// ---- POUs/err.TcPOU
FUNCTION_BLOCK err
VAR_INPUT
	enter : BOOL;
END_VAR
VAR_OUTPUT
END_VAR
VAR
	i:INT;
	step:INT:=0;
	pulse_timer:TON;
	retry_timer:TON;
	has_err:BOOL;
	has_power_not_ready:BOOL;
	has_other_error:BOOL;
	all_powered:BOOL;
	backoff_move : ARRAY[1..7] OF MC_MoveRelative;
	backoff_exec : ARRAY[1..7] OF BOOL;
	backoff_distance : ARRAY[1..7] OF LREAL;
	backoff_attempts : ARRAY[1..7] OF UINT;
	backoff_blocked : BOOL;
	backoff_needed : BOOL;
	backoff_finished : BOOL;
	backoff_error : BOOL;
	backoff_disabled : BOOL;
	power_not_ready_errid : UDINT := 16#00004650;
END_VAR

(* 
Error recovery state:
  - disable external setpoint generation and keep estop hold active
  - if the only active power error is 16#00004650, recover by cycling MC_Power.Enable
  - other errors still use MC_Reset
  - leave _err only after errors are gone and all axes are powered again
*)

has_err := FALSE;
has_power_not_ready := FALSE;
has_other_error := FALSE;
all_powered := TRUE;

FOR i:=1 TO 7 DO
	IF NOT G.power_output[i].Done THEN
		all_powered := FALSE;
	END_IF

	IF G.axis[i].Status.Error OR G.axis[i].Status.DriveDeviceError OR G.power_output[i].Error OR G.reset_output[i].Error THEN
		has_err := TRUE;

		IF (G.power_output[i].Error AND (G.power_output[i].ErrorID = power_not_ready_errid))
		   OR (G.axis[i].Status.Error AND (G.axis[i].Status.ErrorID = power_not_ready_errid)) THEN
			has_power_not_ready := TRUE;
		END_IF

		IF (G.axis[i].Status.Error AND (G.axis[i].Status.ErrorID <> power_not_ready_errid))
		   OR G.axis[i].Status.DriveDeviceError
		   OR G.reset_output[i].Error
		   OR (G.power_output[i].Error AND (G.power_output[i].ErrorID <> power_not_ready_errid)) THEN
			has_other_error := TRUE;
		END_IF
	END_IF
END_FOR

G.estop_hold_req := TRUE;
IF enter THEN
	FOR i:=1 TO 7 DO
		backoff_attempts[i] := 0;
		backoff_exec[i] := FALSE;
		G.err_backoff_failed[i] := FALSE;
		G.err_backoff_active[i] := FALSE;
	END_FOR
END_IF
FOR i:=1 TO 7 DO
	backoff_move[i](Axis:=G.axis[i], Execute:=backoff_exec[i],
		Distance:=backoff_distance[i], Velocity:=G.err_backoff_velocity,
		Acceleration:=G.err_backoff_acc, Deceleration:=G.err_backoff_acc);
END_FOR
backoff_blocked := FALSE;
backoff_needed := FALSE;
IF G.self_check_done AND ((step = 1) OR (step = 3) OR (step = 11)) AND NOT has_err AND all_powered THEN
	backoff_disabled := TRUE;
	FOR i:=1 TO 7 DO
		IF ((i = 1) OR (i = 3) OR (i = 5) OR (i = 6)) AND G.axis[i].Status.DriveLimitActive
			AND G.SetPointGenDisable[i].Enabled THEN backoff_disabled := FALSE; END_IF
	END_FOR
	IF NOT backoff_disabled THEN
		FOR i:=1 TO 7 DO
			G.SetPointGenEnable[i].Execute := FALSE;
			G.SetPointGenDisable[i].Execute := TRUE;
		END_FOR
		RETURN;
	END_IF
	FOR i:=1 TO 7 DO
		IF ((i = 1) OR (i = 3) OR (i = 5) OR (i = 6)) AND G.axis[i].Status.DriveLimitActive THEN
			backoff_blocked := TRUE;
			IF backoff_attempts[i] < G.recovery_max_retries THEN
				IF G.axis[i].NcToPlc.ActPos - G.leftlimit[i] <=
					G.leftlimit[i] + G.rslimit_distance[i] - G.axis[i].NcToPlc.ActPos THEN
					backoff_distance[i] := G.err_backoff_distance;
				ELSE
					backoff_distance[i] := -G.err_backoff_distance;
				END_IF
				backoff_attempts[i] := backoff_attempts[i] + 1;
				backoff_exec[i] := TRUE;
				G.err_backoff_active[i] := TRUE;
				backoff_needed := TRUE;
			ELSE
				G.err_backoff_failed[i] := TRUE;
			END_IF
		END_IF
	END_FOR
	IF backoff_needed THEN step := 20; END_IF
END_IF
IF step = 20 THEN
	backoff_finished := TRUE;
	backoff_error := has_err;
	FOR i:=1 TO 7 DO
		G.SetPointGenEnable[i].Execute := FALSE;
		G.SetPointGenDisable[i].Execute := TRUE;
		IF G.err_backoff_active[i] THEN
			IF backoff_move[i].Error OR backoff_move[i].CommandAborted THEN
				backoff_error := TRUE;
			ELSIF NOT backoff_move[i].Done THEN
				backoff_finished := FALSE;
			END_IF
		END_IF
	END_FOR
	IF backoff_error OR backoff_finished THEN
		FOR i:=1 TO 7 DO
			backoff_exec[i] := FALSE;
			G.err_backoff_active[i] := FALSE;
		END_FOR
		// 重置流程提供下降沿；仍压限位时按本次进入err的剩余次数再退离。
		step := 0;
	END_IF
	RETURN;
END_IF

CASE step OF
0:
	FOR i:=1 TO 7 DO
		G.SetPointGenEnable[i].Execute := FALSE;
		G.SetPointGenDisable[i].Execute := TRUE;
		G.axis_Reset[i].Execute := FALSE;
	END_FOR
	pulse_timer(IN:=FALSE);
	retry_timer(IN:=FALSE);
	step := 1;

1:
	FOR i:=1 TO 7 DO
		G.SetPointGenDisable[i].Execute := FALSE;
	END_FOR

	IF (NOT has_err) AND all_powered AND NOT backoff_blocked THEN
		step := 0;
		G.gen_state := _clear_err;
		RETURN;
	END_IF

	IF NOT has_err THEN
		FOR i:=1 TO 7 DO
			G.axis_Reset[i].Execute := FALSE;
			G.power_[i].Enable := FALSE;
		END_FOR
		pulse_timer(IN:=TRUE, PT:=T#200MS);
		step := 10;
		RETURN;
	END_IF

	IF has_power_not_ready AND NOT has_other_error THEN
		pulse_timer(IN:=TRUE, PT:=T#200MS);
		retry_timer(IN:=FALSE);
		step := 10;
		RETURN;
	END_IF

	FOR i:=1 TO 7 DO
		IF G.axis[i].Status.Error OR G.axis[i].Status.DriveDeviceError OR G.power_output[i].Error OR G.reset_output[i].Error THEN
			G.axis_Reset[i].Execute := TRUE;
		END_IF
	END_FOR
	pulse_timer(IN:=TRUE, PT:=T#200MS);
	step := 2;

2:
	pulse_timer(IN:=TRUE);
	IF pulse_timer.Q THEN
		FOR i:=1 TO 7 DO
			G.axis_Reset[i].Execute := FALSE;
		END_FOR
		pulse_timer(IN:=FALSE);
		retry_timer(IN:=TRUE, PT:=T#2S);
		step := 3;
	END_IF

3:
	retry_timer(IN:=TRUE);

	IF (NOT has_err) AND all_powered AND NOT backoff_blocked THEN
		retry_timer(IN:=FALSE);
		step := 0;
		G.gen_state := _clear_err;
		RETURN;
	END_IF

	IF retry_timer.Q THEN
		retry_timer(IN:=FALSE);
		step := 1;
	END_IF

10:
	FOR i:=1 TO 7 DO
		IF (G.power_output[i].Error AND (G.power_output[i].ErrorID = power_not_ready_errid))
		   OR (G.axis[i].Status.Error AND (G.axis[i].Status.ErrorID = power_not_ready_errid))
		   OR G.axis[i].Status.DriveDeviceError THEN
			G.power_[i].Enable := FALSE;
			G.axis_Reset[i].Execute := TRUE;
		ELSE
			G.power_[i].Enable := TRUE;
			G.axis_Reset[i].Execute := FALSE;
		END_IF
	END_FOR

	pulse_timer(IN:=TRUE, PT:=T#200MS);
	IF pulse_timer.Q THEN
		pulse_timer(IN:=FALSE);
		FOR i:=1 TO 7 DO
			G.axis_Reset[i].Execute := FALSE;
			G.power_[i].Enable := TRUE;
		END_FOR
		retry_timer(IN:=TRUE, PT:=T#3S);
		step := 11;
	END_IF

11:
	FOR i:=1 TO 7 DO
		G.power_[i].Enable := TRUE;
	END_FOR

	retry_timer(IN:=TRUE);

	IF (NOT has_err) AND all_powered AND NOT backoff_blocked THEN
		retry_timer(IN:=FALSE);
		step := 0;
		G.gen_state := _clear_err;
		RETURN;
	END_IF

	IF has_err THEN
		retry_timer(IN:=FALSE);
		step := 1;
		RETURN;
	END_IF

	IF retry_timer.Q THEN
		retry_timer(IN:=FALSE);
		step := 1;
	END_IF
END_CASE

END_FUNCTION_BLOCK

// ---- POUs/reset.TcPOU
FUNCTION_BLOCK reset
VAR_INPUT
END_VAR
VAR_OUTPUT
END_VAR
VAR
	i:INT;
	step:INT:=0;
	reset_timer:TON;
	all_done:BOOL;
END_VAR

(*
FUNCTION_BLOCK: reset
功能说明:
  故障复位流程：对错误轴发出 MC_Reset 清错请求，清错后回到 _init；若错误仍在则转入 _err。

状态机(step):
  0) 预处理：拉低 Execute 形成上升沿；同时请求禁用外部给定模式(避免复位期间被 refer 干预)
  1) 触发复位：对 7 轴发出 MC_Reset.Execute=TRUE，并启动超时计时器
  2) 等待：Done/Error/错误已清除 或超时则收尾并决定跳转(_init/_err)
*)

CASE step OF
0:
	// 预处理：确保后续有上升沿，同时在复位阶段禁用外部给定
	FOR i:=1 TO 7 DO 
		G.axis_Reset[i].Execute := FALSE;
		G.SetPointGenEnable[i].Execute := FALSE;
		G.SetPointGenDisable[i].Execute := TRUE;
	END_FOR
	reset_timer(IN:=FALSE);
	step := 1;

1:
	// 触发复位：Execute 保持 TRUE 直到下个阶段读取 Done/Error
	FOR i:=1 TO 7 DO 
		G.axis_Reset[i].Execute := TRUE;
		// 禁用请求只需要上升沿，避免每周期重复触发
		G.SetPointGenDisable[i].Execute := FALSE;
	END_FOR
	reset_timer(IN:=TRUE, PT:=T#3S);
	step := 2;

2:
	// 等待复位完成（或超时保护）
	reset_timer(IN:=TRUE);
	all_done := TRUE;
	FOR i:=1 TO 7 DO
		IF NOT (G.reset_output[i].Done OR G.reset_output[i].Error OR NOT G.axis[i].Status.Error) THEN 
			all_done := FALSE; 
			EXIT;
		END_IF
	END_FOR
   
	IF all_done OR reset_timer.Q THEN
		// 收尾：撤销 Execute，复位计时器复位，然后返回 init
		FOR i:=1 TO 7 DO 
			G.axis_Reset[i].Execute := FALSE;
		END_FOR
		reset_timer(IN:=FALSE);
		step := 0;

		// 复位结束后，错误已清除才允许回到 _init；否则进入 _err(避免 init/reset 无限循环)
		FOR i:=1 TO 7 DO
			IF G.axis[i].Status.Error OR G.power_output[i].Error OR G.reset_output[i].Error THEN
				G.gen_state := _err;
				RETURN;
			END_IF
		END_FOR
		G.gen_state := _init;
	END_IF
END_CASE

END_FUNCTION_BLOCK

// ---- POUs/SelfCheck.TcPOU
 FUNCTION_BLOCK SelfCheck
VAR_INPUT
    init_target_from_left : ARRAY[1..7] OF LREAL;  // 左限位寻参后回到的工作位（距左限位）
END_VAR
VAR
    i : INT;
    stu : ARRAY[1..7] OF INT; // 0:WaitDisable, 1:StartScan, 2:ScanMonitor, 3:WaitStop, 4:ResetTrigger, 5:WaitReset, 55:RepowerPulse, 56:RepowerWait, 6:SyncWait, 7:SetPosStart, 71:SetPosWait, 72:BackoffDelay, 8:BackoffMove, 10:Done
    fb_move_abs : ARRAY[1..7] OF MC_MoveAbsolute;
    fb_move_vel : ARRAY[1..7] OF MC_MoveVelocity;
    fb_stop     : ARRAY[1..7] OF MC_Stop;
    fb_set_pos  : ARRAY[1..7] OF MC_SetPosition;
    // fb_set_blocked is a function, no instantiation needed
    power_not_ready_errid : UDINT := 16#00004650;
    vel_scan : LREAL := 40.0;   // 寻参逼近速度，>0（单位随轴：mm/s 或 deg/s
    vel_back : LREAL := 40.0;   // 回退速度，>0（单位随轴：mm/s 或 deg/s）

    target_axes : ARRAY[1..7] OF BOOL:= [TRUE,FALSE,TRUE,FALSE,TRUE,TRUE,FALSE];	// 目标轴（平移轴）
    stagger_delay : ARRAY[1..7] OF TIME := [T#3s,T#0ms,T#2s,T#0ms,T#1s,T#0ms,T#0ms];
    scan_stagger_delay : ARRAY[1..7] OF TIME := [T#0ms,T#0ms,T#300ms,T#0ms,T#600ms,T#900ms,T#0ms];
    scan_stagger_timer : ARRAY[1..7] OF TON;
    stagger_started : BOOL := FALSE;
    
    all_done : BOOL;
    all_reach_limit : BOOL;
    
    // 日志触发 (示例)
	Execute: INT;
    
    // 调试变量，用于排查回退距离问题
    debug_limit_pos : ARRAY[1..7] OF LREAL;
    debug_init_target_pos : ARRAY[1..7] OF LREAL;
    scan_start_pos : ARRAY[1..7] OF LREAL;
    
    // 动作控制中间变量，防止多重调用
    mv_vel_exec : ARRAY[1..7] OF BOOL;
    mv_vel_vel  : ARRAY[1..7] OF LREAL;
    mv_abs_exec : ARRAY[1..7] OF BOOL;
    mv_abs_pos : ARRAY[1..7] OF LREAL;
    mv_abs_vel  : ARRAY[1..7] OF LREAL;
    drive_limit_stop : ARRAY[1..7] OF BOOL; // TRUE=电子限位触发路径，等待停止及 Power 状态稳定
    set_pos_exec : ARRAY[1..7] OF BOOL;
    
    // 延时计时器
    wait_timer : ARRAY[1..7] OF TON;
    power_pulse_timer : ARRAY[1..7] OF TON;
    power_wait_timer : ARRAY[1..7] OF TON;
    stagger_timer : TON;
END_VAR

(*
FUNCTION_BLOCK: SelfCheck
功能说明:
  上电自检/寻参流程（负向低速逼近左限位 + 顺序回退），用于建立各轴相对坐标系零点并消除进入外部给定模式前的 SetPos/ActPos 偏差。

自检流程:
  1) 对 target_axes[]包括的平移轴：禁用外部给定（SetPointGenDisable），反向低速逼近左限位并记录 G.leftlimit[]
  2) 对旋转轴（轴2/4/7）：禁用外部给定后，直接 MC_MoveAbsolute 到绝对位置 0
  3) 停止与清错：MC_Stop 平滑停止；若出现故障则 MC_Reset 清错
  4) 目标轴回退：按 seq_order[] 依次 MC_SetPosition(ActPos→SetPos) → MC_MoveAbsolute 回退 → 以回退终点刷新 init_pos[]
  5) 全轴完成后：同步相对坐标变量并切换到 _handle
*)

// 统计：目标轴是否全部进入同步等待阶段（stu>=6）
IF G.selfcheck_reset_req THEN
	G.startup_loading_ready := FALSE;
    FOR i:=1 TO 7 DO
        stu[i] := 0;
        mv_vel_exec[i] := FALSE;
        mv_vel_vel[i] := 0.0;
        mv_abs_exec[i] := FALSE;
        mv_abs_pos[i] := 0.0;
        mv_abs_vel[i] := 0.0;
        drive_limit_stop[i] := FALSE;
        set_pos_exec[i] := FALSE;
        debug_limit_pos[i] := 0.0;
        debug_init_target_pos[i] := 0.0;
        scan_start_pos[i] := 0.0;
        G.selfcheck_stu[i] := 0;
        wait_timer[i](IN:=FALSE);
        scan_stagger_timer[i](IN:=FALSE);
        power_pulse_timer[i](IN:=FALSE);
        power_wait_timer[i](IN:=FALSE);
        G.SetPointGenDisable[i](Axis:=G.axis[i], Execute:=FALSE);
        G.axis_Reset[i](Axis:=G.axis[i], Execute:=FALSE);
        fb_move_vel[i](Axis:=G.axis[i], Execute:=FALSE);
        fb_move_abs[i](Axis:=G.axis[i], Execute:=FALSE);
        fb_stop[i](Axis:=G.axis[i], Execute:=FALSE);
        fb_set_pos[i](Axis:=G.axis[i], Execute:=FALSE);
    END_FOR
    stagger_started := FALSE;
    stagger_timer(IN:=FALSE);
    G.selfcheck_all_reach_limit := FALSE;
    G.axis4_fwd_req := FALSE;
    G.axis4_rev_req := FALSE;
    G.axis4_manual_busy := FALSE;
    G.axis4_manual_done := FALSE;
    G.axis4_manual_error := FALSE;
    G.axis4_manual_error_id := 0;
    G.selfcheck_reset_req := FALSE;
END_IF

// selfcheck 期间固定初始化电缸5，避免阶段切换引入额外切换值。
G.cylinder5_value := 2000;
G.cylinder5_cmd := 2000;
G.cylinder5_press_req := FALSE;

all_reach_limit := TRUE;
FOR i:=1 TO 7 DO
    IF target_axes[i] AND ((stu[i] < 6) OR (NOT G.power_output[i].Done)) THEN
        all_reach_limit := FALSE;
        EXIT;
    END_IF
END_FOR

// 统计：目标轴是否全部处于上电使能状态（避免在 SetPosition 时单轴卡顿）

G.selfcheck_all_reach_limit := all_reach_limit;
stagger_timer(IN:=stagger_started, PT:=T#10s);

FOR i:=1 TO 7 DO
    // 初始化本周期的控制变量

    mv_vel_exec[i] := FALSE;
    mv_abs_exec[i] := FALSE;

    fb_stop[i](Axis:=G.axis[i]);
    IF target_axes[i] THEN
        
        CASE stu[i] OF
        0: // 步骤0：禁用外部给定，避免寻参阶段被外部指令干预
            G.SetPointGenDisable[i](Axis:=G.axis[i], Execute:=TRUE);
            IF G.power_output[i].Done AND (G.SetPointGenDisable[i].Done OR NOT G.SetPointGenDisable[i].Enabled) THEN 
                G.SetPointGenDisable[i](Axis:=G.axis[i], Execute:=FALSE);
                stu[i] := 1;
            END_IF
            
        1: // 错开启动，避免多轴同时加速导致电流竞争触发跟随误差
            IF i = 1 THEN
                G.cylinder1_value := 1000;
                G.cylinder2_value := 10;
				G.cylinder3_value := 1000;
				G.cylinder4_value := 10;
            END_IF

            scan_stagger_timer[i](IN:=TRUE, PT:=scan_stagger_delay[i]);
            IF scan_stagger_timer[i].Q OR scan_stagger_delay[i] = T#0ms THEN
                scan_stagger_timer[i](IN:=FALSE);
                scan_start_pos[i] := G.axis[i].NcToPlc.ActPos;
                drive_limit_stop[i] := FALSE;
                mv_vel_vel[i] := vel_scan;
                mv_vel_exec[i] := TRUE;
                stu[i] := 2;
            END_IF
            
        2:  // 步骤2：监控逼近过程（到限位/堵转判据）
            mv_vel_vel[i] := vel_scan;
            mv_vel_exec[i] := TRUE;
            
            // 电子限位优先；100ms 堵转判据保留为开关或驱动状态失效时的后备保护。
            wait_timer[i](
                IN:= (fb_move_vel[i].Busy
                      AND ABS(G.axis[i].NcToPlc.ActVelo) < 0.5
                      AND (
                          (ABS(G.axis[i].NcToPlc.SetVelo) > 5.0)
                          OR (
                              (ABS(G.axis[i].NcToPlc.SetVelo) < 0.5)
                              AND (ABS(G.axis[i].NcToPlc.ActPos - scan_start_pos[i]) > 1.0)
                          )
                      )),
                PT:= T#100ms
            );
            IF G.axis[i].Status.DriveLimitActive THEN
                // 记录左限位（绝对坐标）
                G.leftlimit[i] := G.axis[i].NcToPlc.ActPos;

                // 立即撤销 MoveVelocity，并在轴状态完全失效前发送受控停止。
                // 现场确认 16#4650 来自 MoveVelocity/MC_Power 就绪链路，而不是 MC_Stop。
                mv_vel_exec[i] := FALSE;
                drive_limit_stop[i] := TRUE;
                wait_timer[i](IN:=FALSE);
                fb_stop[i](
                    Axis:=G.axis[i],
                    Deceleration:=500,
                    Jerk:=1000,
                    Execute:=TRUE
                );
                stu[i] := 3;

            ELSIF fb_move_vel[i].Error OR wait_timer[i].Q THEN
                // 电子限位失效时的后备路径：记录堵转位置并由 MC_Stop 主动停止。
                G.leftlimit[i] := G.axis[i].NcToPlc.ActPos;
                mv_vel_exec[i] := FALSE;
                drive_limit_stop[i] := FALSE;
                fb_stop[i](
                    Axis:=G.axis[i], 
                    Deceleration:=500, 
                    Jerk:=1000, 
                    Execute:=TRUE
                );
                stu[i] := 3;
            END_IF
            
        3: // 步骤3：等待停止完成（以 ActVelo 作为停稳判据）
            IF ABS(G.axis[i].NcToPlc.ActVelo) < 1.0 THEN
                fb_stop[i](Axis:=G.axis[i], Execute:=FALSE);

                IF drive_limit_stop[i] THEN
                    // DriveLimitActive 后 Disabled/Power 状态存在延迟，等待其稳定后再决定恢复路径。
                    wait_timer[i](IN:=TRUE, PT:=T#300ms);
                    IF wait_timer[i].Q THEN
                        wait_timer[i](IN:=FALSE);

                        IF G.axis[i].Status.Error
                           OR (G.power_output[i].Error AND (G.power_output[i].ErrorID <> power_not_ready_errid))
                        THEN
                            drive_limit_stop[i] := FALSE;
                            stu[i] := 4;
                        ELSIF G.power_output[i].Done AND NOT G.power_output[i].Error THEN
                            drive_limit_stop[i] := FALSE;
                            stu[i] := 6;
                        ELSE
                            // 电子限位导致的 16#4650/Power not ready 通过 MC_Power 下降沿重新初始化。
                            power_pulse_timer[i](IN:=FALSE);
                            power_wait_timer[i](IN:=FALSE);
                            stu[i] := 55;
                        END_IF
                    END_IF
                ELSE
                    wait_timer[i](IN:=FALSE);
                    IF G.axis[i].Status.Error THEN
                        stu[i] := 4;
                    ELSIF G.power_output[i].Done AND NOT G.power_output[i].Error THEN
                        stu[i] := 6;
                    ELSE
                        power_pulse_timer[i](IN:=FALSE);
                        power_wait_timer[i](IN:=FALSE);
                        stu[i] := 55;
                    END_IF
                END_IF
            ELSE
                wait_timer[i](IN:=FALSE);
            END_IF
            
        4: // 步骤4：触发错误清除（通常为限位/跟随相关故障）
            G.axis_Reset[i](Axis:=G.axis[i], Execute:=FALSE);
            G.axis_Reset[i](Axis:=G.axis[i], Execute:=TRUE);
            // 触发后立即进入等待，避免同周期重复触发
            stu[i] := 5;
            
        5: // 步骤5：等待错误清除完成
            G.axis_Reset[i](Axis:=G.axis[i]);
            power_pulse_timer[i](IN:=FALSE);
            power_wait_timer[i](IN:=FALSE);
            
            IF G.axis_Reset[i].Done OR NOT G.axis[i].Status.Error THEN
                G.axis_Reset[i](Axis:=G.axis[i], Execute:=FALSE);
                // 进入同步等待：后续统一进行 SetPosition + 回退
                IF G.power_output[i].Done THEN
                    stu[i] := 6;
                ELSE
                    power_pulse_timer[i](IN:=FALSE);
                    power_wait_timer[i](IN:=FALSE);
                    IF i = 6 THEN
                        stagger_started := FALSE;
                        stagger_timer(IN:=FALSE);
                    END_IF
                    stu[i] := 55;
                END_IF
            ELSIF G.axis_Reset[i].Error THEN
                // 复位失败，尝试重试
                G.axis_Reset[i](Axis:=G.axis[i], Execute:=FALSE);
                stu[i] := 4;
            END_IF
        55: // RepowerPulse: 关闭 MC_Power Enable 一个脉冲，让轴重新初始化
            G.power_[i].Enable := FALSE;
            power_pulse_timer[i](IN:=TRUE, PT:=T#200ms);
            IF power_pulse_timer[i].Q THEN
                power_pulse_timer[i](IN:=FALSE);
                G.power_[i].Enable := TRUE;
                stu[i] := 56;
            END_IF

        56: // RepowerWait: 等待 MC_Power 重新就绪
            G.power_[i].Enable := TRUE;
            power_wait_timer[i](IN:=TRUE, PT:=T#3s);
            IF G.power_output[i].Done AND NOT G.power_output[i].Error THEN
                power_wait_timer[i](IN:=FALSE);
                drive_limit_stop[i] := FALSE;
                stu[i] := 6;
            ELSIF power_wait_timer[i].Q THEN
                // 超时仍未就绪，重试
                power_wait_timer[i](IN:=FALSE);
                power_pulse_timer[i](IN:=FALSE);
                stu[i] := 55;
            END_IF
		6: // 步骤6：同步等待（全部目标轴都到达后，同时放行回退）
            IF all_reach_limit AND G.power_output[i].Done THEN
                stu[i] := 7;
            ELSIF NOT G.power_output[i].Done THEN
                power_pulse_timer[i](IN:=FALSE);
                power_wait_timer[i](IN:=FALSE);
                IF i = 6 THEN
                    stagger_started := FALSE;
                    stagger_timer(IN:=FALSE);
                END_IF
                stu[i] := 55;
            END_IF
            
        7: // 步骤7：同步 SetPos=ActPos，避免进入回退/外部给定时产生突跳
            IF NOT G.power_output[i].Done THEN
                set_pos_exec[i] := FALSE;
                fb_set_pos[i](Axis:=G.axis[i], Execute:=FALSE);
                power_pulse_timer[i](IN:=FALSE);
                power_wait_timer[i](IN:=FALSE);
                IF i = 6 THEN
                    stagger_started := FALSE;
                    stagger_timer(IN:=FALSE);
                END_IF
                stu[i] := 55;
            ELSE
				set_pos_exec[i] := TRUE;
				fb_set_pos[i](
					Axis:=G.axis[i],
					Position:=G.axis[i].NcToPlc.ActPos,
					Mode:=FALSE,
					Execute:=set_pos_exec[i]
				);
				stu[i] := 71;
            END_IF

        71: // 步骤71：等待位置同步完成，然后启动回退
            fb_set_pos[i](Axis:=G.axis[i], Execute:=set_pos_exec[i]);
            
            IF NOT G.power_output[i].Done THEN
                set_pos_exec[i] := FALSE;
                fb_set_pos[i](Axis:=G.axis[i], Execute:=FALSE);
                power_pulse_timer[i](IN:=FALSE);
                power_wait_timer[i](IN:=FALSE);
                IF i = 6 THEN
                    stagger_started := FALSE;
                    stagger_timer(IN:=FALSE);
                END_IF
                stu[i] := 55;
            ELSIF fb_set_pos[i].Done THEN
				set_pos_exec[i] := FALSE;
                fb_set_pos[i](Axis:=G.axis[i], Execute:=FALSE);
                
               
                // 启动绝对回退（目标=左限位绝对坐标 + 回退距离）
                debug_limit_pos[i] := G.leftlimit[i];
                debug_init_target_pos[i] := G.leftlimit[i] + init_target_from_left[i];
                
                mv_abs_pos[i] := debug_init_target_pos[i];
                mv_abs_vel[i] := vel_back;
                mv_abs_exec[i] := FALSE;
                wait_timer[i](IN:=FALSE);
                
                stu[i] := 72;
             
            ELSIF fb_set_pos[i].Error THEN
                // 如果 SetPosition 失败，尝试重试复位
				set_pos_exec[i] := FALSE;
                fb_set_pos[i](Axis:=G.axis[i], Execute:=FALSE);
                IF G.power_output[i].Error THEN
                    power_pulse_timer[i](IN:=FALSE);
                    power_wait_timer[i](IN:=FALSE);
                    IF i = 6 THEN
                        stagger_started := FALSE;
                        stagger_timer(IN:=FALSE);
                    END_IF
                    stu[i] := 55;
                ELSE
                    stu[i] := 4;
                END_IF
            END_IF

        72: // 步骤72：轴6先发起并确认回退，其他目标轴按 stagger_delay 依次放行
            mv_abs_pos[i] := debug_init_target_pos[i];
            mv_abs_vel[i] := vel_back;
            mv_abs_exec[i] := FALSE;

            wait_timer[i](IN:=FALSE);
            IF i = 6 THEN
                IF NOT G.power_output[i].Done THEN
                    power_pulse_timer[i](IN:=FALSE);
                    power_wait_timer[i](IN:=FALSE);
                    stagger_started := FALSE;
                    stagger_timer(IN:=FALSE);
                    stu[i] := 55;
                ELSE
                    mv_abs_exec[i] := TRUE;
                    IF fb_move_abs[i].Busy OR fb_move_abs[i].Done OR (ABS(G.axis[i].NcToPlc.ActVelo) > 0.5) THEN
                        IF NOT stagger_started THEN
                            stagger_started := TRUE;
                            stagger_timer(IN:=FALSE);
                        END_IF
                        stu[i] := 8;
                    END_IF
                END_IF
            ELSIF stagger_started AND (stagger_timer.ET >= stagger_delay[i]) THEN
                IF G.power_output[i].Done THEN
                    mv_abs_exec[i] := TRUE;
                    stu[i] := 8;
                ELSE
                    power_pulse_timer[i](IN:=FALSE);
                    power_wait_timer[i](IN:=FALSE);
                    stu[i] := 55;
                END_IF
            END_IF
            
        8: // 步骤8：等待回退完成
            mv_abs_pos[i] := debug_init_target_pos[i];
            mv_abs_vel[i] := vel_back;
            mv_abs_exec[i] := TRUE;
            
            IF fb_move_abs[i].Done THEN
                mv_abs_exec[i] := FALSE;
                stu[i] := 10; // 完成
			ELSIF fb_move_abs[i].Error OR fb_move_abs[i].CommandAborted THEN
				mv_abs_exec[i] := FALSE;
				IF G.power_output[i].Error THEN
					// Power 层面出了问题，先重新上电
					power_pulse_timer[i](IN:=FALSE);
					power_wait_timer[i](IN:=FALSE);
                    IF i = 6 THEN
                        stagger_started := FALSE;
                        stagger_timer(IN:=FALSE);
                    END_IF
					stu[i] := 55;
				ELSE
					stu[i] := 4;
				END_IF
			END_IF
            
        10: // 完成：以回退终点作为新的相对零点（刷新 init_pos）
            G.init_pos[i] := G.axis[i].NcToPlc.ActPos;
        END_CASE
    ELSE
        // 轴4保持当前位置；轴2/7回到绝对位置0。
        IF i = 4 THEN
            CASE stu[i] OF
            0:
                G.SetPointGenDisable[i](Axis:=G.axis[i], Execute:=TRUE);
                IF G.power_output[i].Done AND (G.SetPointGenDisable[i].Done OR NOT G.SetPointGenDisable[i].Enabled) THEN
                    G.SetPointGenDisable[i](Axis:=G.axis[i], Execute:=FALSE);
                    stu[i] := 10;
                END_IF
            10:
                G.init_pos[i] := G.axis[i].NcToPlc.ActPos;
            END_CASE
        ELSE
        CASE stu[i] OF
        0: // 禁用外部给定，避免与绝对定位冲突
            G.SetPointGenDisable[i](Axis:=G.axis[i], Execute:=TRUE);
            IF G.power_output[i].Done AND (G.SetPointGenDisable[i].Done OR NOT G.SetPointGenDisable[i].Enabled) THEN
                G.SetPointGenDisable[i](Axis:=G.axis[i], Execute:=FALSE);
                stu[i] := 1;
            END_IF

        1: // 启动绝对定位到 0
            mv_abs_pos[i] := 0.0;
            mv_abs_vel[i] := vel_back;
            mv_abs_exec[i] := TRUE;
            stu[i] := 2;

        2: // 等待到位
            mv_abs_pos[i] := 0.0;
            mv_abs_vel[i] := vel_back;
            mv_abs_exec[i] := TRUE;

            IF fb_move_abs[i].Done
               OR (NOT fb_move_abs[i].Busy AND ABS(G.axis[i].NcToPlc.ActPos - mv_abs_pos[i]) < 0.01)
            THEN
                mv_abs_exec[i] := FALSE;
                stu[i] := 10;
            ELSIF fb_move_abs[i].Error OR fb_move_abs[i].CommandAborted THEN
                mv_abs_exec[i] := FALSE;
                stu[i] := 4;
            END_IF

        4: // 触发复位清错
            G.axis_Reset[i](Axis:=G.axis[i], Execute:=FALSE);
            G.axis_Reset[i](Axis:=G.axis[i], Execute:=TRUE);
            stu[i] := 5;

        5: // 等待复位完成后重试定位
            G.axis_Reset[i](Axis:=G.axis[i]);
            IF G.axis_Reset[i].Done OR NOT G.axis[i].Status.Error THEN
                G.axis_Reset[i](Axis:=G.axis[i], Execute:=FALSE);
                stu[i] := 1;
            ELSIF G.axis_Reset[i].Error THEN
                G.axis_Reset[i](Axis:=G.axis[i], Execute:=FALSE);
                stu[i] := 4;
            END_IF
        END_CASE
        END_IF
    END_IF
    
    // 统一调用运动控制功能块 (在每个周期末尾)
    fb_move_vel[i](
        Axis:=G.axis[i],
        Execute:=mv_vel_exec[i],
        Velocity:=mv_vel_vel[i],
        Acceleration:=50,
        Deceleration:=100,
        Jerk:=100,
        Direction:=MC_Direction.MC_Negative_Direction
    );
    fb_move_abs[i](
        Axis:=G.axis[i], 
        Position:=mv_abs_pos[i], 
        Velocity:=mv_abs_vel[i], 
        Acceleration:=100, 
        Deceleration:=100, 
        Jerk:=100,
        Execute:=mv_abs_exec[i]
    );
	G.selfcheck_stu[i] := stu[i];
END_FOR

// 全轴完成判定（所有轴 stu=10）
all_done := TRUE;
FOR i:=1 TO 7 DO
    IF stu[i] <> 10 THEN
        all_done := FALSE;
        EXIT;
    END_IF
END_FOR

IF all_done THEN
	G.cylinder1_value := 1000;
	G.cylinder2_value := 150;
	G.cylinder3_value := 1000;
	G.cylinder4_value := 150;
    G.self_check_done := TRUE;
	G.startup_loading_ready := TRUE;
    G.handle_reinit_req := TRUE;
    FOR i:=1 TO 7 DO
        // 旋转轴已回到绝对零位，参考坐标必须同样采用绝对零点。
        // 不能保留 init 阶段采集的自检前角度，否则相对 0 会重新指向旧位置。
        IF NOT target_axes[i] AND i <> 4 THEN
            G.init_pos[i] := 0.0;
        ELSIF i = 4 THEN
            G.init_pos[i] := G.axis[i].NcToPlc.ActPos;
        END_IF
        // 统一刷新相对坐标/参考，避免切换到 handle 后出现参考突变
        G.Act_pos[i] := G.axis[i].NcToPlc.ActPos - G.init_pos[i];
        G.act_pos_from_left[i] := G.axis[i].NcToPlc.ActPos - G.leftlimit[i];
        G.refer[i] := G.Act_pos[i];
        G.ref_slow[i] := G.Act_pos[i];
        G.act_h[i] := G.Act_pos[i];
        G.act_hf[i] := G.Act_pos[i];
        G.refer_from_left[i] := G.act_pos_from_left[i];
    END_FOR
    G.gen_state := _handle;
END_IF

END_FUNCTION_BLOCK

// ---- POUs/ArmManual.TcPOU
FUNCTION_BLOCK ArmManual
VAR
	i : INT;
	req_dir : SINT;
	cmd_velocity : LREAL;
	cmd_acc : LREAL;
	cmd_dec : LREAL;
	cmd_jerk : LREAL;
	allow_jog : BOOL;

	// 每轴独立状态：0=空闲，10=点动中，20=停止中，30=换向停止中
	axis_state : ARRAY[1..5] OF INT := [0,0,0,0,0];
	current_dir : ARRAY[1..5] OF SINT := [0,0,0,0,0];
	pending_dir : ARRAY[1..5] OF SINT := [0,0,0,0,0];
	move_exec : ARRAY[1..5] OF BOOL := [FALSE,FALSE,FALSE,FALSE,FALSE];
	stop_exec : ARRAY[1..5] OF BOOL := [FALSE,FALSE,FALSE,FALSE,FALSE];
	reset_exec : ARRAY[1..5] OF BOOL := [FALSE,FALSE,FALSE,FALSE,FALSE];
	move_direction : ARRAY[1..5] OF MC_Direction;

	fb_power : ARRAY[1..5] OF MC_Power;
	fb_reset : ARRAY[1..5] OF MC_Reset;
	fb_move_vel : ARRAY[1..5] OF MC_MoveVelocity;
	fb_stop : ARRAY[1..5] OF MC_Stop;
END_VAR

FOR i:=1 TO 5 DO
	// 定位臂轴独立刷新，不影响介入机器人 G.axis[1..7] 主链路
	G.arm_axis[i]();
	G.arm_act_pos[i] := G.arm_axis[i].NcToPlc.ActPos;
	G.arm_act_vel[i] := G.arm_axis[i].NcToPlc.ActVelo;
	IF G.host_comm_timeout OR NOT G.arm_manual_enable THEN
		// 主机看门狗超时或总使能关闭后均不继承单轴上电和点动请求。
		// 该保护独立于原 7 轴状态机，避免上位机异常退出后定位臂继续带电。
		G.arm_manual_enable := FALSE;
		G.arm_enable_req[i] := FALSE;
		G.arm_jog_pos_req[i] := FALSE;
		G.arm_jog_neg_req[i] := FALSE;
	END_IF

	cmd_velocity := G.arm_jog_velocity[i];
	IF cmd_velocity <= 0.0 THEN
		cmd_velocity := 5.0;
	END_IF
	cmd_acc := G.arm_jog_acc[i];
	IF cmd_acc <= 0.0 THEN
		cmd_acc := 50.0;
	END_IF
	cmd_dec := G.arm_jog_dec[i];
	IF cmd_dec <= 0.0 THEN
		cmd_dec := 50.0;
	END_IF
	cmd_jerk := G.arm_jog_jerk[i];
	IF cmd_jerk <= 0.0 THEN
		cmd_jerk := 500.0;
	END_IF

	fb_power[i](
		Axis:=G.arm_axis[i],
		Enable:=G.arm_manual_enable AND G.arm_enable_req[i],
		Enable_Positive:=TRUE,
		Enable_Negative:=TRUE
	);
	G.arm_power_output[i].Done := fb_power[i].Status;
	G.arm_power_output[i].Busy := fb_power[i].Busy;
	G.arm_power_output[i].Active := fb_power[i].Active;
	G.arm_power_output[i].Error := fb_power[i].Error;
	G.arm_power_output[i].ErrorID := fb_power[i].ErrorID;

	IF G.arm_reset_req[i] AND NOT reset_exec[i] THEN
		IF G.arm_curve_owned OR G.arm_cjog_owned THEN
			IF G.arm_curve_owned THEN G.arm_curve_cancel := TRUE; END_IF
		ELSE
		reset_exec[i] := TRUE;
		move_exec[i] := FALSE;
		stop_exec[i] := TRUE;
		axis_state[i] := 20;
		current_dir[i] := 0;
		END_IF
	END_IF

	// 复位请求先等待 MC_Stop 完成，避免清错瞬间释放尚未停止的旧运动命令。
	fb_reset[i](Axis:=G.arm_axis[i], Execute:=reset_exec[i] AND (axis_state[i] = 0));
	G.arm_reset_output[i].Done := fb_reset[i].Done;
	G.arm_reset_output[i].Busy := fb_reset[i].Busy OR reset_exec[i];
	G.arm_reset_output[i].Active := FALSE;
	G.arm_reset_output[i].Error := fb_reset[i].Error;
	G.arm_reset_output[i].ErrorID := fb_reset[i].ErrorID;
	IF reset_exec[i] AND (fb_reset[i].Done OR fb_reset[i].Error) THEN
		IF fb_reset[i].Done AND NOT G.arm_axis[i].Status.Error THEN
			G.arm_motion_error[i] := FALSE;
			G.arm_motion_error_id[i] := 0;
			G.arm_motion_done[i] := TRUE;
		ELSIF fb_reset[i].Error THEN
			G.arm_motion_error[i] := TRUE;
			G.arm_motion_error_id[i] := fb_reset[i].ErrorID;
		END_IF
		reset_exec[i] := FALSE;
		G.arm_reset_req[i] := FALSE;
	END_IF

	G.arm_cmd_conflict[i] := G.arm_jog_pos_req[i] AND G.arm_jog_neg_req[i];
	IF G.arm_cmd_conflict[i] THEN
		req_dir := 0;
	ELSIF G.arm_jog_pos_req[i] THEN
		req_dir := 1;
	ELSIF G.arm_jog_neg_req[i] THEN
		req_dir := -1;
	ELSE
		req_dir := 0;
	END_IF

	allow_jog := G.arm_manual_enable
		AND NOT G.arm_curve_owned
		AND NOT G.arm_cjog_owned
		AND G.arm_power_output[i].Done
		AND NOT reset_exec[i]
		AND NOT G.arm_cmd_conflict[i]
		AND NOT G.arm_axis[i].Status.Error
		AND NOT G.arm_power_output[i].Error
		AND NOT G.arm_reset_output[i].Error;
	IF NOT allow_jog THEN
		req_dir := 0;
	END_IF

	IF fb_move_vel[i].Error THEN
		G.arm_motion_error[i] := TRUE;
		G.arm_motion_error_id[i] := fb_move_vel[i].ErrorID;
		move_exec[i] := FALSE;
		stop_exec[i] := FALSE;
		current_dir[i] := 0;
		axis_state[i] := 0;
	ELSIF fb_stop[i].Error THEN
		G.arm_motion_error[i] := TRUE;
		G.arm_motion_error_id[i] := fb_stop[i].ErrorID;
		move_exec[i] := FALSE;
		stop_exec[i] := FALSE;
		current_dir[i] := 0;
		axis_state[i] := 0;
	END_IF

	CASE axis_state[i] OF
	0: // 空闲，等待新的正/反点动命令
		move_exec[i] := FALSE;
		stop_exec[i] := FALSE;
		current_dir[i] := 0;
		pending_dir[i] := 0;
		IF req_dir <> 0 THEN
			IF req_dir > 0 THEN
				move_direction[i] := MC_Direction.MC_Positive_Direction;
			ELSE
				move_direction[i] := MC_Direction.MC_Negative_Direction;
			END_IF
			move_exec[i] := TRUE;
			current_dir[i] := req_dir;
			G.arm_motion_done[i] := FALSE;
			G.arm_motion_error[i] := FALSE;
			G.arm_motion_error_id[i] := 0;
			axis_state[i] := 10;
		END_IF

	10: // 点动中：松开即停，方向变化先停稳再反向启动
		stop_exec[i] := FALSE;
		IF req_dir = 0 THEN
			move_exec[i] := FALSE;
			stop_exec[i] := TRUE;
			current_dir[i] := 0;
			axis_state[i] := 20;
		ELSIF req_dir <> current_dir[i] THEN
			move_exec[i] := FALSE;
			stop_exec[i] := TRUE;
			pending_dir[i] := req_dir;
			current_dir[i] := 0;
			axis_state[i] := 30;
		ELSE
			move_exec[i] := TRUE;
		END_IF

	20: // 常规停止
		move_exec[i] := FALSE;
		stop_exec[i] := TRUE;
		IF fb_stop[i].Done OR ((ABS(G.arm_act_vel[i]) < 0.01) AND NOT fb_stop[i].Busy) THEN
			stop_exec[i] := FALSE;
			G.arm_motion_done[i] := TRUE;
			axis_state[i] := 0;
		END_IF

	30: // 换向停止，停稳后仍保持新方向按钮才重新启动
		move_exec[i] := FALSE;
		stop_exec[i] := TRUE;
		IF fb_stop[i].Done OR ((ABS(G.arm_act_vel[i]) < 0.01) AND NOT fb_stop[i].Busy) THEN
			stop_exec[i] := FALSE;
			IF (pending_dir[i] <> 0) AND (req_dir = pending_dir[i]) THEN
				IF pending_dir[i] > 0 THEN
					move_direction[i] := MC_Direction.MC_Positive_Direction;
				ELSE
					move_direction[i] := MC_Direction.MC_Negative_Direction;
				END_IF
				move_exec[i] := TRUE;
				current_dir[i] := pending_dir[i];
				pending_dir[i] := 0;
				G.arm_motion_done[i] := FALSE;
				G.arm_motion_error[i] := FALSE;
				G.arm_motion_error_id[i] := 0;
				axis_state[i] := 10;
			ELSE
				pending_dir[i] := 0;
				G.arm_motion_done[i] := TRUE;
				axis_state[i] := 0;
			END_IF
		END_IF

	ELSE
		move_exec[i] := FALSE;
		stop_exec[i] := FALSE;
		current_dir[i] := 0;
		pending_dir[i] := 0;
		axis_state[i] := 0;
	END_CASE

	fb_move_vel[i](
		Axis:=G.arm_axis[i],
		Execute:=move_exec[i],
		Velocity:=cmd_velocity,
		Acceleration:=cmd_acc,
		Deceleration:=cmd_dec,
		Jerk:=cmd_jerk,
		Direction:=move_direction[i]
	);

	fb_stop[i](
		Axis:=G.arm_axis[i],
		Execute:=stop_exec[i],
		Deceleration:=cmd_dec,
		Jerk:=cmd_jerk
	);

	IF G.arm_axis[i].Status.Error THEN
		G.arm_motion_error[i] := TRUE;
		IF G.arm_power_output[i].Error THEN
			G.arm_motion_error_id[i] := G.arm_power_output[i].ErrorID;
		ELSIF G.arm_reset_output[i].Error THEN
			G.arm_motion_error_id[i] := G.arm_reset_output[i].ErrorID;
		ELSE
			G.arm_motion_error_id[i] := 0;
		END_IF
	END_IF

	G.arm_cmd_dir[i] := current_dir[i];
	G.arm_motion_busy[i] := (axis_state[i] <> 0) OR fb_move_vel[i].Busy OR fb_stop[i].Busy OR reset_exec[i];
END_FOR

END_FUNCTION_BLOCK

// ---- POUs/ArmCartesian.TcPOU
FUNCTION_BLOCK ArmCartesian
VAR
    stage : INT;
    i : INT;
    k : INT;
    curve : ARRAY[0..16] OF LREAL;
    incoming : ARRAY[0..16] OF LREAL;
    p : ARRAY[1..5] OF LREAL;
    v : ARRAY[1..5] OF LREAL;
    a : ARRAY[1..5] OF LREAL;
    dir : ARRAY[1..5] OF DINT;
    velocity_limit : ARRAY[1..5] OF LREAL;
    acceleration_limit : ARRAY[1..5] OF LREAL;
    deceleration_limit : ARRAY[1..5] OF LREAL;
    jerk_limit : ARRAY[1..5] OF LREAL;
    elapsed : LREAL;
    phase_elapsed : LREAL;
    cycle_seconds : LREAL;
    segment_seconds : LREAL;
    u : LREAL;
    path_progress : LREAL;
    ds : LREAL;
    dds : LREAL;
    delta : LREAL;
    bend : LREAL;
    slope_bound : LREAL;
    allowed : BOOL;
    drive_ready : BOOL;
    all_enabled : BOOL;
    all_disabled : BOOL;
    all_stopped : BOOL;
    all_released : BOOL;
    arrived : BOOL;
    reject_error : UDINT;
    last_heartbeat : UDINT;
    heartbeat_age : LREAL;
    finish_state : UDINT;
    fb_enable : ARRAY[1..5] OF MC_ExtSetPointGenEnable;
    fb_disable : ARRAY[1..5] OF MC_ExtSetPointGenDisable;
    fb_stop : ARRAY[1..5] OF MC_Stop;
END_VAR

// 定位臂归零保留原1ms曲线接口，第16项必须为0。
cycle_seconds := UDINT_TO_LREAL(TwinCAT_SystemInfoVarList._TaskInfo[1].CycleTime) * 0.0000001;
IF TwinCAT_SystemInfoVarList._TaskInfo[1].FirstCycle THEN
    G.arm_curve_ack := G.arm_curve_request;
    G.arm_curve_cancel := TRUE;
    G.arm_curve_owned := FALSE;
    G.arm_curve_state := 0;
    G.arm_curve_error := 0;
    stage := 0;
END_IF
IF G.arm_curve_heartbeat <> last_heartbeat THEN
    last_heartbeat := G.arm_curve_heartbeat;
    heartbeat_age := 0;
ELSE
    heartbeat_age := heartbeat_age + cycle_seconds;
END_IF

drive_ready := G.arm_manual_enable AND NOT G.host_comm_timeout AND NOT G.estop_hold_req
    AND (ABS(cycle_seconds - 0.001) < 0.00000001);
FOR i := 1 TO 5 DO
    drive_ready := drive_ready AND G.arm_power_output[i].Done AND G.arm_enable_req[i]
        AND NOT G.arm_axis[i].Status.Error AND NOT G.arm_reset_req[i]
        AND NOT G.arm_jog_pos_req[i] AND NOT G.arm_jog_neg_req[i];
END_FOR
allowed := drive_ready AND (heartbeat_age < 0.5);

IF G.arm_curve_request <> G.arm_curve_ack THEN
    IF stage >= 40 THEN
        // 停止中的迟到请求只确认接收，不重新启动运动。
        IF G.arm_curve_error = 0 THEN G.arm_curve_error := 2001; END_IF
        finish_state := 4;
        G.arm_curve_cancel := TRUE;
        G.arm_curve_ack := G.arm_curve_request;
    ELSE
        reject_error := 0;
        FOR k := 0 TO 16 DO
            incoming[k] := G.arm_curve_data[k];
            IF NOT ((incoming[k] >= -100000.0) AND (incoming[k] <= 100000.0)) THEN
                reject_error := 2002;
            END_IF
        END_FOR
        IF (incoming[15] < 0.02) OR (incoming[15] > 120.0)
            OR (incoming[16] <> 0.0) THEN
            reject_error := 2002;
        END_IF
        IF NOT allowed OR G.arm_curve_cancel THEN reject_error := 2003; END_IF
        IF (stage <> 0) AND (reject_error = 0) THEN reject_error := 2001; END_IF
        IF G.arm_cjog_owned THEN reject_error := 2001; END_IF

        IF reject_error = 0 THEN
            FOR i := 1 TO 5 DO
                IF NOT ((G.arm_jog_velocity[i] > 0) AND (G.arm_jog_velocity[i] <= 10000))
                    OR NOT ((G.arm_jog_acc[i] > 0) AND (G.arm_jog_acc[i] <= 10000))
                    OR NOT ((G.arm_jog_dec[i] > 0) AND (G.arm_jog_dec[i] <= 10000))
                    OR NOT ((G.arm_jog_jerk[i] > 0) AND (G.arm_jog_jerk[i] <= 10000)) THEN
                    reject_error := 2002;
                END_IF
            END_FOR
        END_IF
        IF reject_error = 0 THEN
            FOR i := 1 TO 5 DO
                delta := incoming[i+4] - incoming[i-1];
                segment_seconds := incoming[15];
                    bend := incoming[i+9];
                    IF ABS(bend) > ABS(delta)/4.0+0.000000001 THEN reject_error := 2002; END_IF
                    slope_bound := ABS(delta)+4.0*ABS(bend);
                    IF (1.875*slope_bound/segment_seconds > G.arm_jog_velocity[i]+0.0000001)
                        OR ((6.0*slope_bound+28.125*ABS(bend))/(segment_seconds*segment_seconds)
                            > G.arm_jog_acc[i]+0.0000001) THEN
                        reject_error := 2005;
                    END_IF

            END_FOR
            IF (MIN(incoming[4],incoming[9]) < -60.0)
                OR (MAX(incoming[4],incoming[9]) > 60.0) THEN reject_error := 2006; END_IF
        END_IF
        IF reject_error = 0 THEN
            FOR i := 1 TO 5 DO
                // 负载下反馈会波动，启动只依据忙状态，不用速度或起点偏差判停稳。
                IF G.arm_motion_busy[i] THEN
                    reject_error := 2004;
                END_IF
            END_FOR
        END_IF

        IF reject_error = 0 THEN
                FOR k := 0 TO 16 DO curve[k] := incoming[k]; END_FOR
                FOR i := 1 TO 5 DO
                    p[i] := curve[i-1];
                    v[i] := 0;
                    a[i] := 0;
                    dir[i] := 0;
                    IF curve[i+4] > p[i] THEN dir[i] := 1; END_IF
                    IF curve[i+4] < p[i] THEN dir[i] := -1; END_IF
                    velocity_limit[i] := G.arm_jog_velocity[i];
                    acceleration_limit[i] := G.arm_jog_acc[i];
                    deceleration_limit[i] := G.arm_jog_dec[i];
                    jerk_limit[i] := G.arm_jog_jerk[i];
                END_FOR
                G.arm_curve_owned := TRUE;
                stage := 10;
                elapsed := 0;
                phase_elapsed := 0;
                finish_state := 2;
                G.arm_curve_progress := 0;
            G.arm_curve_error := 0;
            G.arm_curve_state := 1;
        ELSE
            IF G.arm_curve_error = 0 THEN G.arm_curve_error := reject_error; END_IF
            G.arm_curve_cancel := TRUE;
            finish_state := 4;
            IF stage > 0 THEN
                stage := 40;
                phase_elapsed := 0;
            END_IF
        END_IF
        // 先锁存归零曲线，再确认序号。
        G.arm_curve_ack := G.arm_curve_request;
    END_IF
END_IF

IF (stage > 0) AND (stage < 40) THEN
    IF G.arm_curve_cancel OR NOT allowed THEN
        finish_state := 3;
        IF NOT allowed THEN
            IF G.arm_curve_error = 0 THEN G.arm_curve_error := 2003; END_IF
            finish_state := 4; G.arm_curve_cancel := TRUE;
        END_IF
        stage := 40;
        phase_elapsed := 0;
    END_IF
END_IF
IF stage > 0 THEN phase_elapsed := phase_elapsed + cycle_seconds; END_IF
IF (stage = 10 OR stage = 30) AND (phase_elapsed > 2.0) THEN
    IF G.arm_curve_error = 0 THEN G.arm_curve_error := 2007; END_IF
    G.arm_curve_cancel := TRUE;
    finish_state := 4;
    stage := 40;
END_IF

IF stage = 20 THEN
    u := MIN(1.0, elapsed/curve[15]);
    path_progress := u*u*u*(10.0+u*(-15.0+6.0*u));
    ds := 30.0*u*u*(1.0-u)*(1.0-u)/curve[15];
    dds := 60.0*u*(1.0-u)*(1.0-2.0*u)/(curve[15]*curve[15]);
    FOR i := 1 TO 5 DO
        delta := curve[i+4]-curve[i-1];
            bend := curve[i+9];
            p[i] := curve[i-1]+path_progress*delta+4.0*path_progress*(1.0-path_progress)*bend;
            v[i] := (delta+4.0*(1.0-2.0*path_progress)*bend)*ds;
            a[i] := (delta+4.0*(1.0-2.0*path_progress)*bend)*dds-8.0*bend*ds*ds;
        IF (ABS(v[i]) > velocity_limit[i]+0.000001)
            OR (ABS(a[i]) > acceleration_limit[i]+0.000001)
            OR NOT ((G.arm_act_pos[i]-p[i] >= -1.0) AND (G.arm_act_pos[i]-p[i] <= 1.0)) THEN
            IF G.arm_curve_error = 0 THEN G.arm_curve_error := 2008; END_IF
            G.arm_curve_cancel := TRUE;
            finish_state := 4;
            stage := 40;
        END_IF
    END_FOR
    G.arm_curve_progress := u;
    elapsed := elapsed+cycle_seconds;
    IF (u >= 1.0) AND (stage = 20) THEN
        stage := 30;
        phase_elapsed := 0;
    END_IF
END_IF

all_enabled := TRUE;
all_disabled := TRUE;
all_stopped := TRUE;
all_released := TRUE;
arrived := TRUE;
FOR i := 1 TO 5 DO
    // 归零沿用原外部设定点发生器握手。
    IF G.arm_curve_owned THEN
        MC_ExtSetPointGenFeed(Axis:=G.arm_axis[i], Position:=p[i],
            Velocity:=v[i], Acceleration:=a[i], Direction:=dir[i]);
    END_IF
    fb_enable[i](Axis:=G.arm_axis[i], Execute:=(stage=10),
        Position:=curve[i+4], PositionType:=POSITIONTYPE_ABSOLUTE);
    fb_disable[i](Axis:=G.arm_axis[i], Execute:=(stage=40));
    fb_stop[i](Axis:=G.arm_axis[i], Execute:=(stage=50) AND NOT G.arm_axis[i].Status.Error,
        Deceleration:=deceleration_limit[i], Jerk:=jerk_limit[i]);
    all_enabled := all_enabled AND fb_enable[i].Enabled;
    // 与末端点动相同，错误轴和功能块错误不阻塞所有权释放。
    all_disabled := all_disabled AND (fb_disable[i].Done OR fb_disable[i].Error OR G.arm_axis[i].Status.Error);
    all_stopped := all_stopped AND (fb_stop[i].Done OR fb_stop[i].Error OR G.arm_axis[i].Status.Error);
    all_released := all_released AND NOT fb_stop[i].Busy;
    arrived := arrived AND (ABS(G.arm_act_pos[i]-curve[i+4]) <= 0.05)
        AND (ABS(G.arm_act_vel[i]) <= 0.1);
    IF G.arm_curve_owned AND (fb_enable[i].Error OR fb_disable[i].Error OR fb_stop[i].Error) THEN
        G.arm_curve_cancel := TRUE;
        IF G.arm_curve_error = 0 THEN
            IF fb_enable[i].Error THEN G.arm_curve_error := fb_enable[i].ErrorID;
            ELSIF fb_disable[i].Error THEN G.arm_curve_error := fb_disable[i].ErrorID;
            ELSIF fb_stop[i].Error THEN G.arm_curve_error := fb_stop[i].ErrorID; END_IF
        END_IF
        finish_state := 4;
        IF stage < 40 THEN stage := 40; END_IF
    END_IF
END_FOR

CASE stage OF
10:
    IF all_enabled THEN stage := 20; elapsed := 0; phase_elapsed := 0; END_IF
30:
    IF arrived AND (phase_elapsed >= 2.0*cycle_seconds) THEN stage := 40; END_IF
40:
    IF all_disabled THEN
        IF finish_state = 2 THEN stage := 60; ELSE stage := 50; END_IF
    END_IF
50:
    IF all_stopped THEN stage := 60; END_IF
60:
    IF all_released THEN
        G.arm_curve_owned := FALSE;
        G.arm_curve_state := finish_state;
        stage := 0;
    END_IF
END_CASE
IF G.arm_curve_error <> 0 THEN
    G.arm_curve_state := 4;
END_IF

END_FUNCTION_BLOCK

// ---- POUs/ArmCartJog.TcPOU
FUNCTION_BLOCK ArmCartJog
VAR CONSTANT
    ALIVE_TIMEOUT : LREAL := 0.5; // 秒
    ENABLE_TIMEOUT : LREAL := 2.0;
END_VAR
VAR
    stage : INT;
    i : INT;
    cycle_seconds : LREAL;
    alive_age : LREAL;
    enable_age : LREAL;
    last_alive : UDINT;
    request_valid : BOOL;
    held : BOOL;
    drive_ready : BOOL;
    fault_stop : BOOL;
    all_enabled, all_disabled, all_stopped, all_released : BOOL;
    zero_cycles : INT;
    dir_feed : ARRAY[1..5] OF DINT;
    gen : ArmCartJogGen;
    fb_enable : ARRAY[1..5] OF MC_ExtSetPointGenEnable;
    fb_disable : ARRAY[1..5] OF MC_ExtSetPointGenDisable;
    fb_stop : ARRAY[1..5] OF MC_Stop;
END_VAR

cycle_seconds := UDINT_TO_LREAL(TwinCAT_SystemInfoVarList._TaskInfo[1].CycleTime)*0.0000001;
IF TwinCAT_SystemInfoVarList._TaskInfo[1].FirstCycle THEN
    stage := 0;
    G.arm_cjog_owned := FALSE;
    G.arm_cjog_state := 0;
    G.arm_cjog_error := 0;
    G.arm_cjog_limited := FALSE;
    G.arm_cjog_path_speed := 0;
END_IF
IF G.arm_cjog_alive <> last_alive THEN
    last_alive := G.arm_cjog_alive;
    alive_age := 0;
ELSE
    alive_age := alive_age+cycle_seconds;
END_IF
// ADS请求只在此边界校验；mode=0是正常松开。
request_valid := (G.arm_cjog_mode >= 1) AND (G.arm_cjog_mode <= 5)
    AND ((G.arm_cjog_dir = -1) OR (G.arm_cjog_dir = 1))
    AND (G.arm_cjog_speed > 0) AND (G.arm_cjog_speed <= 100);
held := request_valid AND (alive_age < ALIVE_TIMEOUT);
IF (G.arm_cjog_mode <> 0) AND NOT request_valid AND (G.arm_cjog_error = 0) THEN G.arm_cjog_error := 3001; END_IF
// 与ArmCartesian的驱动就绪表达式逐项一致。
drive_ready := G.arm_manual_enable AND NOT G.host_comm_timeout AND NOT G.estop_hold_req
    AND (ABS(cycle_seconds-0.001) < 0.00000001);
FOR i := 1 TO 5 DO
    drive_ready := drive_ready AND G.arm_power_output[i].Done AND G.arm_enable_req[i]
        AND NOT G.arm_axis[i].Status.Error AND NOT G.arm_reset_req[i]
        AND NOT G.arm_jog_pos_req[i] AND NOT G.arm_jog_neg_req[i];
END_FOR
IF (stage = 0) AND held AND NOT G.arm_curve_owned
    AND (G.arm_curve_request = G.arm_curve_ack) THEN
    IF NOT drive_ready THEN
        IF G.arm_cjog_error = 0 THEN G.arm_cjog_error := 3002; END_IF
    ELSE
        gen(start:=TRUE, held:=FALSE, mode:=G.arm_cjog_mode, dir:=G.arm_cjog_dir,
            speed:=G.arm_cjog_speed, seed:=G.arm_act_pos, cycle_dt:=cycle_seconds);
        FOR i := 1 TO 5 DO dir_feed[i] := 1; END_FOR
        G.arm_cjog_error := 0;
        G.arm_cjog_owned := TRUE;
        fault_stop := FALSE;
        enable_age := 0;
        zero_cycles := 0;
        stage := 10;
    END_IF
END_IF
IF (stage = 10 OR stage = 25) AND NOT drive_ready THEN
    IF G.arm_cjog_error = 0 THEN G.arm_cjog_error := 3002; END_IF
    fault_stop := TRUE;
    stage := 40;
END_IF
IF stage = 10 THEN
    enable_age := enable_age+cycle_seconds;
    IF enable_age > ENABLE_TIMEOUT THEN
        IF G.arm_cjog_error = 0 THEN G.arm_cjog_error := 3003; END_IF
        fault_stop := TRUE;
        stage := 40;
    END_IF
END_IF
IF stage = 25 THEN
    gen(start:=FALSE, held:=held, mode:=G.arm_cjog_mode, dir:=G.arm_cjog_dir,
        speed:=G.arm_cjog_speed, seed:=gen.p, cycle_dt:=cycle_seconds);
    IF (gen.path_speed = 0) AND NOT held THEN
        zero_cycles := zero_cycles+1;
    ELSE
        zero_cycles := 0;
    END_IF
    IF zero_cycles >= 2 THEN stage := 40; END_IF
END_IF
all_enabled := TRUE; all_disabled := TRUE; all_stopped := TRUE; all_released := TRUE;
FOR i := 1 TO 5 DO
    IF gen.v[i] > 0 THEN dir_feed[i] := 1; END_IF
    IF gen.v[i] < 0 THEN dir_feed[i] := -1; END_IF
    IF G.arm_cjog_owned AND (stage = 10 OR stage = 25) THEN
        MC_ExtSetPointGenFeed(Axis:=G.arm_axis[i], Position:=gen.p[i],
            Velocity:=gen.v[i], Acceleration:=gen.a[i], Direction:=dir_feed[i]);
    END_IF
    fb_enable[i](Axis:=G.arm_axis[i], Execute:=(stage=10),
        Position:=gen.p[i], PositionType:=POSITIONTYPE_ABSOLUTE);
    fb_disable[i](Axis:=G.arm_axis[i], Execute:=(stage=40));
    fb_stop[i](Axis:=G.arm_axis[i], Execute:=(stage=50) AND NOT G.arm_axis[i].Status.Error,
        Deceleration:=G.arm_jog_dec[i], Jerk:=G.arm_jog_jerk[i]);
    all_enabled := all_enabled AND fb_enable[i].Enabled;
    // 错误轴交回NC复位；停用或停止报错也必须走完释放。
    all_disabled := all_disabled AND (fb_disable[i].Done OR fb_disable[i].Error OR G.arm_axis[i].Status.Error);
    all_stopped := all_stopped AND (fb_stop[i].Done OR fb_stop[i].Error OR G.arm_axis[i].Status.Error);
    all_released := all_released AND NOT fb_stop[i].Busy;
    IF G.arm_cjog_owned AND (fb_enable[i].Error OR fb_disable[i].Error OR fb_stop[i].Error) THEN
        IF G.arm_cjog_error = 0 THEN
            IF fb_enable[i].Error THEN G.arm_cjog_error := fb_enable[i].ErrorID;
            ELSIF fb_disable[i].Error THEN G.arm_cjog_error := fb_disable[i].ErrorID;
            ELSIF fb_stop[i].Error THEN G.arm_cjog_error := fb_stop[i].ErrorID; END_IF
        END_IF
        fault_stop := TRUE;
        IF stage < 40 THEN stage := 40; END_IF
    END_IF
END_FOR
CASE stage OF
10:
    IF all_enabled THEN stage := 25; END_IF
40:
    IF all_disabled THEN
        IF fault_stop THEN stage := 50; ELSE stage := 60; END_IF
    END_IF
50:
    IF all_stopped THEN stage := 60; END_IF
60:
    IF all_released THEN G.arm_cjog_owned := FALSE; stage := 0; END_IF
END_CASE
CASE stage OF
0: G.arm_cjog_state := 0;
10: G.arm_cjog_state := 1;
25:
    IF gen.target_speed > 0 THEN G.arm_cjog_state := 2;
    ELSE G.arm_cjog_state := 3; END_IF
40,50,60: G.arm_cjog_state := 4;
END_CASE
G.arm_cjog_limited := gen.limited;
G.arm_cjog_path_speed := gen.path_speed;

END_FUNCTION_BLOCK

// ---- POUs/ArmCartJogGen.TcPOU
FUNCTION_BLOCK ArmCartJogGen
VAR_INPUT
    start : BOOL;
    held : BOOL;
    mode : INT;
    dir : INT;
    speed : LREAL;
    seed : ARRAY[1..5] OF LREAL;
    cycle_dt : LREAL;
END_VAR
VAR_OUTPUT
    p : ARRAY[1..5] OF LREAL;
    v : ARRAY[1..5] OF LREAL;
    a : ARRAY[1..5] OF LREAL;
    path_speed : LREAL;
    target_speed : LREAL;
    limited : BOOL;
END_VAR
VAR CONSTANT
    PI : LREAL := 3.14159265358979323846;
    RAD : LREAL := PI / 180.0;
    L1 : LREAL := 200.0; // 毫米，取自kinematics.h
    L2 : LREAL := 180.0;
    TOOL_LATERAL_OFFSET_MM : LREAL := 456.3;
    TOOL_LENGTH_MM : LREAL := 554.5;
    T_ACC : LREAL := 1.0; // 秒
    T_DEC : LREAL := 0.5;
    INITIAL_BRANCH : INT := 1;
    BISECTION_COUNT : INT := 12;
    JOINT_VCAP : ARRAY[1..5] OF LREAL := [24,30,30,30,30]; // 毫米/秒、度/秒
END_VAR
VAR
    anchor : ARRAY[1..5] OF LREAL;
    position_before, velocity_before : ARRAY[1..5] OF LREAL;
    path_v, path_v_previous, v0, v1, tau, sigma : LREAL;
    duration : LREAL := T_ACC;
    wx, wy : LREAL;
    psi0, d0x, d0y, tcp0x, tcp0y : LREAL;
    latched_mode, latched_dir : INT;
    branch : INT := INITIAL_BRANCH;
    reanchor, trial_ok : BOOL;
    i, j : INT;
    u, delta_sigma_des, delta_sigma, lower_step, upper_step : LREAL;
    best_step, trial_step, axis_sign, signed_path, ex, ey : LREAL;
    candidate_wx, candidate_wy, best_wx, best_wy : LREAL;
    candidate_radius, candidate_cosine, candidate_elbow : LREAL;
    candidate_azimuth, azimuth_denominator : LREAL;
    candidate_q2, candidate_q3, candidate_q4 : LREAL;
    candidate_psi : LREAL;
    best_q2, best_q3, best_q4, branch_q3 : LREAL;
END_VAR

// 输入速度采用平滑曲线，路径增量用相邻周期速度的梯形积分。
reanchor := start;
IF start THEN
    p := seed;
    FOR i := 1 TO 5 DO v[i] := 0; a[i] := 0; END_FOR
    path_v := 0; v0 := 0; v1 := 0; tau := 0; duration := T_ACC;
    latched_mode := mode; latched_dir := dir;
END_IF
position_before := p; velocity_before := v; path_v_previous := path_v;
target_speed := 0;
IF held AND (mode = latched_mode) AND (dir = latched_dir) THEN target_speed := speed; END_IF
IF target_speed <> v1 THEN
    v0 := path_v; v1 := target_speed;
    IF v1 > v0 THEN duration := T_ACC; ELSE duration := T_DEC; END_IF
    tau := 0;
END_IF
IF NOT start THEN tau := tau + cycle_dt; END_IF
u := MIN(1.0, tau / duration);
path_v := v0 + (v1-v0)*(3.0*u*u-2.0*u*u*u);
// 模式或方向变化在曲线零速点重新锚定。
IF (path_v = 0) AND (v1 = 0) AND held
    AND ((mode <> latched_mode) OR (dir <> latched_dir)) THEN reanchor := TRUE; END_IF
IF reanchor THEN
    anchor := p; latched_mode := mode; latched_dir := dir; sigma := 0;
    branch_q3 := anchor[3];
    WHILE branch_q3 > 180.0 DO branch_q3 := branch_q3-360.0; END_WHILE
    WHILE branch_q3 < -180.0 DO branch_q3 := branch_q3+360.0; END_WHILE
    IF (branch_q3 <> 0.0) AND (branch_q3 <> 180.0) AND (branch_q3 <> -180.0) THEN
        IF branch_q3 < 0 THEN branch := 1; ELSE branch := -1; END_IF
    END_IF
    wx := L1*SIN(anchor[2]*RAD)+L2*SIN((anchor[2]+anchor[3])*RAD+PI);
    wy := -L1*COS(anchor[2]*RAD)-L2*COS((anchor[2]+anchor[3])*RAD+PI);
    psi0 := anchor[2]+anchor[3]+anchor[4];
    d0x := TOOL_LATERAL_OFFSET_MM;
    d0y := -TOOL_LENGTH_MM*COS(anchor[5]*RAD);
    tcp0x := wx+d0x*COS(psi0*RAD)-d0y*SIN(psi0*RAD);
    tcp0y := wy+d0x*SIN(psi0*RAD)+d0y*COS(psi0*RAD);
END_IF
limited := FALSE;
IF start THEN path_speed := 0; target_speed := 0; RETURN; END_IF
delta_sigma_des := 0.5*(path_v_previous+path_v)*cycle_dt;
IF latched_mode = 5 THEN
    // 每周期由偏航累计角和锚定TCP反求腕点，不累加腕点位移。
    best_step := 0; lower_step := 0; upper_step := delta_sigma_des;
    FOR i := 0 TO BISECTION_COUNT DO
        IF i = 0 THEN trial_step := delta_sigma_des;
        ELSE trial_step := (lower_step+upper_step)/2.0; END_IF
        candidate_psi := psi0+latched_dir*(sigma+trial_step);
        candidate_wx := tcp0x-d0x*COS(candidate_psi*RAD)+d0y*SIN(candidate_psi*RAD);
        candidate_wy := tcp0y-d0x*SIN(candidate_psi*RAD)-d0y*COS(candidate_psi*RAD);
        candidate_radius := SQRT(candidate_wx*candidate_wx+candidate_wy*candidate_wy);
        trial_ok := FALSE;
        IF (candidate_radius >= L1-L2) AND (candidate_radius <= L1+L2) THEN
            candidate_cosine := (candidate_radius*candidate_radius-L1*L1-L2*L2)/(2.0*L1*L2);
            IF candidate_cosine > 1.0 THEN candidate_cosine := 1.0;
            ELSIF candidate_cosine < -1.0 THEN candidate_cosine := -1.0; END_IF
            candidate_elbow := branch*ACOS(candidate_cosine);
            azimuth_denominator := -candidate_wy;
            IF azimuth_denominator > 0 THEN candidate_azimuth := ATAN(candidate_wx/azimuth_denominator);
            ELSIF azimuth_denominator < 0 THEN
                IF candidate_wx >= 0 THEN candidate_azimuth := ATAN(candidate_wx/azimuth_denominator)+PI;
                ELSE candidate_azimuth := ATAN(candidate_wx/azimuth_denominator)-PI; END_IF
            ELSE
                IF candidate_wx > 0 THEN candidate_azimuth := PI/2.0;
                ELSE candidate_azimuth := -PI/2.0; END_IF
            END_IF
            candidate_q2 := (candidate_azimuth-ATAN(L2*SIN(candidate_elbow)/(L1+L2*COS(candidate_elbow))))/RAD;
            candidate_q3 := (candidate_elbow-PI)/RAD;
            WHILE candidate_q2-p[2] > 180.0 DO candidate_q2 := candidate_q2-360.0; END_WHILE
            WHILE candidate_q2-p[2] < -180.0 DO candidate_q2 := candidate_q2+360.0; END_WHILE
            WHILE candidate_q3-p[3] > 180.0 DO candidate_q3 := candidate_q3-360.0; END_WHILE
            WHILE candidate_q3-p[3] < -180.0 DO candidate_q3 := candidate_q3+360.0; END_WHILE
            candidate_q4 := anchor[4]+(candidate_psi-psi0)-((candidate_q2+candidate_q3)-(anchor[2]+anchor[3]));
            trial_ok := (ABS(candidate_q2-p[2]) <= JOINT_VCAP[2]*cycle_dt)
                AND (ABS(candidate_q3-p[3]) <= JOINT_VCAP[3]*cycle_dt)
                AND (ABS(candidate_q4-p[4]) <= JOINT_VCAP[4]*cycle_dt);
        END_IF
        IF trial_ok THEN
            lower_step := trial_step; best_step := trial_step;
            best_wx := candidate_wx; best_wy := candidate_wy;
            best_q2 := candidate_q2; best_q3 := candidate_q3; best_q4 := candidate_q4;
            IF i = 0 THEN EXIT; END_IF
        ELSE
            upper_step := trial_step;
        END_IF
    END_FOR
    delta_sigma := best_step;
    IF delta_sigma > 0 THEN
        p[1] := anchor[1]; p[5] := anchor[5];
        p[2] := best_q2; p[3] := best_q3; p[4] := best_q4;
    END_IF
ELSIF latched_mode >= 3 THEN
    // Z正向为轴1减小；俯仰正向为轴5减小。
    IF latched_mode = 3 THEN j := 1;
    ELSIF latched_mode = 4 THEN j := 5;
    ELSE j := 4; END_IF
    delta_sigma := MIN(delta_sigma_des, JOINT_VCAP[j]*cycle_dt);
    signed_path := latched_dir*(sigma+delta_sigma);
    p := anchor;
    axis_sign := -1.0;
    p[j] := anchor[j]+axis_sign*signed_path;
ELSE
    // X/Y试探直线步长；环带与三关节步长共同决定可接受步长。
    IF latched_mode = 1 THEN ex := 1.0; ey := 0.0;
    ELSE ex := 0.0; ey := 1.0; END_IF
    best_step := 0; lower_step := 0; upper_step := delta_sigma_des;
    FOR i := 0 TO BISECTION_COUNT DO
        IF i = 0 THEN trial_step := delta_sigma_des;
        ELSE trial_step := (lower_step+upper_step)/2.0; END_IF
        candidate_wx := wx+latched_dir*trial_step*ex;
        candidate_wy := wy+latched_dir*trial_step*ey;
        candidate_radius := SQRT(candidate_wx*candidate_wx+candidate_wy*candidate_wy);
        trial_ok := FALSE;
        IF (candidate_radius >= L1-L2) AND (candidate_radius <= L1+L2) THEN
            candidate_cosine := (candidate_radius*candidate_radius-L1*L1-L2*L2)/(2.0*L1*L2);
            IF candidate_cosine > 1.0 THEN candidate_cosine := 1.0;
            ELSIF candidate_cosine < -1.0 THEN candidate_cosine := -1.0; END_IF
            candidate_elbow := branch*ACOS(candidate_cosine);
            azimuth_denominator := -candidate_wy;
            IF azimuth_denominator > 0 THEN candidate_azimuth := ATAN(candidate_wx/azimuth_denominator);
            ELSIF azimuth_denominator < 0 THEN
                IF candidate_wx >= 0 THEN candidate_azimuth := ATAN(candidate_wx/azimuth_denominator)+PI;
                ELSE candidate_azimuth := ATAN(candidate_wx/azimuth_denominator)-PI; END_IF
            ELSE
                IF candidate_wx > 0 THEN candidate_azimuth := PI/2.0;
                ELSE candidate_azimuth := -PI/2.0; END_IF
            END_IF
            candidate_q2 := (candidate_azimuth-ATAN(L2*SIN(candidate_elbow)/(L1+L2*COS(candidate_elbow))))/RAD;
            candidate_q3 := (candidate_elbow-PI)/RAD;
            WHILE candidate_q2-p[2] > 180.0 DO candidate_q2 := candidate_q2-360.0; END_WHILE
            WHILE candidate_q2-p[2] < -180.0 DO candidate_q2 := candidate_q2+360.0; END_WHILE
            WHILE candidate_q3-p[3] > 180.0 DO candidate_q3 := candidate_q3-360.0; END_WHILE
            WHILE candidate_q3-p[3] < -180.0 DO candidate_q3 := candidate_q3+360.0; END_WHILE
            candidate_q4 := anchor[4]+(anchor[2]+anchor[3])-(candidate_q2+candidate_q3);
            trial_ok := (ABS(candidate_q2-p[2]) <= JOINT_VCAP[2]*cycle_dt)
                AND (ABS(candidate_q3-p[3]) <= JOINT_VCAP[3]*cycle_dt)
                AND (ABS(candidate_q4-p[4]) <= JOINT_VCAP[4]*cycle_dt);
        END_IF
        IF trial_ok THEN
            lower_step := trial_step; best_step := trial_step;
            best_wx := candidate_wx; best_wy := candidate_wy;
            best_q2 := candidate_q2; best_q3 := candidate_q3; best_q4 := candidate_q4;
            IF i = 0 THEN EXIT; END_IF
        ELSE
            upper_step := trial_step;
        END_IF
    END_FOR
    delta_sigma := best_step;
    IF delta_sigma > 0 THEN
        wx := best_wx; wy := best_wy;
        p[1] := anchor[1]; p[5] := anchor[5];
        p[2] := best_q2; p[3] := best_q3; p[4] := best_q4;
    END_IF
END_IF
sigma := sigma+delta_sigma;
path_speed := delta_sigma/cycle_dt;
limited := delta_sigma < delta_sigma_des;
FOR i := 1 TO 5 DO
    v[i] := (p[i]-position_before[i])/cycle_dt;
    a[i] := (v[i]-velocity_before[i])/cycle_dt;
END_FOR

END_FUNCTION_BLOCK

// ---- POUs/Axis2Sync.TcPOU
FUNCTION_BLOCK Axis2Sync
VAR
	reset_pulse : TON;
	reset_interval : TON;
	reset_execute : BOOL;
	had_axis_error : BOOL;
	fb_power : MC_Power;
	fb_gear : MC_GearIn;
	fb_reset : MC_Reset;
	gear_execute : BOOL := FALSE;
	gear_active : BOOL := FALSE;
	gear_done : BOOL := FALSE;
	gear_failed : BOOL := FALSE;
END_VAR

G.axis2_sync_axis();

G.axis2_sync_error := G.axis2_sync_axis.Status.Error OR G.axis2_sync_axis.Status.DriveDeviceError;
G.axis2_sync_error_id := G.axis2_sync_axis.Status.ErrorID;
IF G.axis2_sync_error THEN
    reset_interval(IN:=TRUE, PT:=G.axis15_reset_interval);
    IF NOT had_axis_error THEN
        reset_execute := TRUE;
    ELSIF reset_interval.Q THEN
        reset_execute := TRUE;
        reset_interval(IN:=FALSE);
    END_IF
	reset_pulse(IN:=reset_execute, PT:=G.axis15_reset_pulse);
	IF reset_pulse.Q THEN reset_execute := FALSE; END_IF
ELSE
	reset_execute := FALSE;
	reset_pulse(IN:=FALSE);
	reset_interval(IN:=FALSE);
	IF had_axis_error THEN
		gear_execute := FALSE;
		gear_active := FALSE;
		gear_done := FALSE;
		gear_failed := FALSE;
	END_IF
END_IF
had_axis_error := G.axis2_sync_error;
fb_reset(
	Axis:=G.axis2_sync_axis,
	Execute:=G.axis_Reset[2].Execute OR reset_execute
);

fb_power(
	Axis:=G.axis2_sync_axis,
	Enable:=G.power_[2].Enable,
	Enable_Positive:=TRUE,
	Enable_Negative:=TRUE
);

IF NOT (G.power_[2].Enable AND G.power_output[2].Done AND fb_power.Status) THEN
	gear_execute := FALSE;
	gear_active := FALSE;
	gear_done := FALSE;
	gear_failed := FALSE;
ELSIF NOT G.axis2_sync_error AND fb_power.Status AND G.power_output[2].Done AND NOT gear_done AND NOT gear_failed AND NOT gear_active
	AND (ABS(G.axis[2].NcToPlc.ActVelo) <= 0.01)
	AND (ABS(G.axis2_sync_axis.NcToPlc.ActVelo) <= 0.01) THEN
	gear_execute := TRUE;
	gear_active := TRUE;
END_IF

fb_gear(
	Master:=G.axis[2],
	Slave:=G.axis2_sync_axis,
	Execute:=gear_execute,
	RatioNumerator:=1.0,
	RatioDenominator:=1,
	Acceleration:=100.0,
	Deceleration:=100.0,
	Jerk:=500.0,
	BufferMode:=MC_Aborting
);

IF fb_gear.InGear THEN
	gear_execute := FALSE;
	gear_active := FALSE;
	gear_done := TRUE;
ELSIF fb_gear.Error OR fb_gear.CommandAborted THEN
	gear_execute := FALSE;
	gear_active := FALSE;
	gear_failed := TRUE;
END_IF

END_FUNCTION_BLOCK

// ---- POUs/InjectorManual.TcPOU
FUNCTION_BLOCK InjectorManual
VAR
	i : INT;
	req_dir : SINT;
	cmd_velocity : LREAL := 180.0;
	cmd_acc : LREAL := 100.0;
	cmd_dec : LREAL := 100.0;
	cmd_jerk : LREAL := 500.0;
	axis_state : ARRAY[1..2] OF INT := [0,0];
	current_dir : ARRAY[1..2] OF SINT := [0,0];
	pending_dir : ARRAY[1..2] OF SINT := [0,0];
	move_exec : ARRAY[1..2] OF BOOL := [FALSE,FALSE];
	stop_exec : ARRAY[1..2] OF BOOL := [FALSE,FALSE];
	move_direction : ARRAY[1..2] OF MC_Direction;
	fb_power : ARRAY[1..2] OF MC_Power;
	fb_move_vel : ARRAY[1..2] OF MC_MoveVelocity;
	fb_stop : ARRAY[1..2] OF MC_Stop;
END_VAR

FOR i:=1 TO 2 DO
	IF G.host_comm_timeout THEN
		G.inject_push_req[i] := FALSE;
		G.inject_pull_req[i] := FALSE;
	END_IF

	fb_power[i](
		Axis:=G.inject_axis[i],
		Enable:=TRUE,
		Enable_Positive:=TRUE,
		Enable_Negative:=TRUE
	);

	IF G.inject_push_req[i] AND NOT G.inject_pull_req[i] THEN
		req_dir := 1;
	ELSIF G.inject_pull_req[i] AND NOT G.inject_push_req[i] THEN
		req_dir := -1;
	ELSE
		req_dir := 0;
	END_IF

	IF axis_state[i] = 0 THEN
		IF req_dir <> 0 THEN
			current_dir[i] := req_dir;
			IF req_dir > 0 THEN
				move_direction[i] := MC_Direction.MC_Positive_Direction;
			ELSE
				move_direction[i] := MC_Direction.MC_Negative_Direction;
			END_IF
			move_exec[i] := TRUE;
			axis_state[i] := 10;
		END_IF
	ELSIF axis_state[i] = 10 THEN
		IF req_dir = current_dir[i] THEN
			move_exec[i] := TRUE;
		ELSIF req_dir <> 0 THEN
			pending_dir[i] := req_dir;
			move_exec[i] := FALSE;
			stop_exec[i] := TRUE;
			current_dir[i] := 0;
			axis_state[i] := 30;
		ELSE
			pending_dir[i] := 0;
			move_exec[i] := FALSE;
			stop_exec[i] := TRUE;
			current_dir[i] := 0;
			axis_state[i] := 20;
		END_IF
	ELSIF axis_state[i] = 20 OR axis_state[i] = 30 THEN
		move_exec[i] := FALSE;
		stop_exec[i] := TRUE;
		IF fb_stop[i].Done OR (ABS(G.inject_axis[i].NcToPlc.ActVelo) <= 0.05) THEN
			stop_exec[i] := FALSE;
			IF axis_state[i] = 30 AND pending_dir[i] <> 0 AND req_dir = pending_dir[i] THEN
				current_dir[i] := pending_dir[i];
				IF current_dir[i] > 0 THEN
					move_direction[i] := MC_Direction.MC_Positive_Direction;
				ELSE
					move_direction[i] := MC_Direction.MC_Negative_Direction;
				END_IF
				move_exec[i] := TRUE;
				pending_dir[i] := 0;
				axis_state[i] := 10;
			ELSE
				current_dir[i] := 0;
				pending_dir[i] := 0;
				axis_state[i] := 0;
			END_IF
		END_IF
	END_IF

	fb_move_vel[i](
		Axis:=G.inject_axis[i],
		Execute:=move_exec[i],
		Velocity:=cmd_velocity,
		Acceleration:=cmd_acc,
		Deceleration:=cmd_dec,
		Jerk:=cmd_jerk,
		Direction:=move_direction[i]
	);
	fb_stop[i](
		Axis:=G.inject_axis[i],
		Execute:=stop_exec[i],
		Deceleration:=cmd_dec,
		Jerk:=cmd_jerk
	);
END_FOR

END_FUNCTION_BLOCK
